(* IEC 61131-3 sources: repolevel_ST_code_completion/dataset/project_code/VisuElements/PRG, 4 files *)

(* ---- MAIN.st ---- *)
PROGRAM MAIN
VAR

END_VAR

(* expand and collapse a node*)
Node();

(* several mouse events *)
MouseEvents();

(* calculate the rotation points for an object *)
Rotation();

(* ---- MouseEvents.st ---- *)
PROGRAM Node
VAR
	xNodeExpand   : BOOL;
	NodeDblClick  : TON;
	tNodeDblClick : TIME := T#500MS; (* the time to wait for the second click *)
	xNodeClick    : BOOL;
	xNodeClickOld : BOOL;
	iNodeState    : INT := 1;
	xNodeSelected : BOOL;
END_VAR

(* This program ellapses/collapses a node, by dozble clicking the first node *)

CASE iNodeState OF

	1: (* first click on the node
		  the first click toggles the xNodeClick variable to true*)
		IF xNodeClick AND NOT xNodeClickOld THEN
			NodeDblClick(IN:=TRUE, PT:=tNodeDblClick);
			iNodeState    := 2;
		END_IF

	2: (* The second click expands respectively collapses the Node *)
		NodeDblClick();
		(* the time for the second click is elapsed*)
		IF NodeDblClick.Q THEN
			NodeDblClick(IN:=FALSE);
			xNodeClick := xNodeClickOld := FALSE;
			iNodeState := 1;
		ELSE
		(* check for the second click,
			when xNodeClick is false, the user has clicked the second time, because xNodeClick is toggled*)
			IF NOT xNodeClick AND xNodeClickOld THEN
				NodeDblClick(IN:=FALSE);
				xNodeExpand := NOT xNodeExpand;
				iNodeState  := 1;
			END_IF
		END_IF
END_CASExNodeClickOld := xNodeClick;

(* ---- Node.st ---- *)
PROGRAM MAIN
VAR

END_VAR

(* expand and collapse a node*)
Node();

(* several mouse events *)
MouseEvents();

(* calculate the rotation points for an object *)
Rotation();

(* ---- Rotation.st ---- *)
PROGRAM MAIN
VAR

END_VAR

(* expand and collapse a node*)
Node();

(* several mouse events *)
MouseEvents();

(* calculate the rotation points for an object *)
Rotation();
